Fanuc KAREL source: KD00034.KL

PROGRAM KD00034
%NOLOCKGROUP
VAR
  I: INTEGER
  J: INTEGER
  B: BOOLEAN
  R: REAL
  S: STRING[80]
BEGIN
  CONDITION[1]:
  WHEN I > 1 DO
    I = 1
  ENDCONDITION
END KD00034
